// System API/DSM/API/bds_dsm_getErrors_DTC
///This function is used to get all DTCs with the specified status.
///
///=======
/// Remarks:
///=======
///    + The |GVL_dsm| is given for usage of defines.
///	
///----------
/// FFI:
///----------
///This API can be used in trusted partitions only. See Freedom from Interference (FFI) concept for more details.
///
///==================================================================		  			===================================================================================================
///Return value    								  									Description
///==================================================================		  			===================================================================================================
///16#0000: BDS_DSM_NO_ERROR_DU16														Got all DTC with specified status.
///16#0004: BDS_DSM_INVALID_PTR_DU16													Invalid Pointer.
///16#0005: BDS_DSM_MASK_ERROR_DU16													Invalid Mask.
///16#0007: BDS_DSM_INVALID_MAX_ERROR_DU16 											Invalid Max number of errors.
///16#0008:BDS_DSM_OVERFLOW_ERROR_DU16													Number of error are more than Max Error. 
///
///==================================================================		   			===================================================================================================
///
///
///=======
///Code Example:
///=======
///============================================================================
///
///PROGRAM DSM
///
///VAR
///
///	mask_s : UINT := BDS_DSM_SET_ACTIVE_ERROR_MASK_DU16;
///
///	startFromBegin_l: BOOL := TRUE;
///
///	maxNum_u16:UINT := 32;
///
///	error_count_u16: UINT;
///
///	dtc_u16: ARRAY [1..32] OF UINT;
///
///	status_u16: UINT;
///
///END_VAR
///
///
///(*Get errors*)
///
///status_u16 := bds_dsm_getErrors(mask_s,startFromBegin_l,maxNum_u16,ADR(error_count_u16),ADR(dtc_u16)); 
///
///IF status_u16 = BDS_DSM_NO_ERROR_DU16 THEN
///
///	(*Number of Errors has been read successfully*)
///
///END_IF
///
///============================================================================
///
{attribute 'external_name' := 'cmp_rts_bds_dsm_getErrors_DTC'}
FUNCTION bds_dsm_getErrors_DTC : UINT
VAR_INPUT
	///The kind of error status can be specified in detail by means of this mask.
	///
	///Possible values:
	///    + BDS_DSM_SET_ACTIVE_ERROR_MASK_DU16 ( 16#18 ) - Fault is active.
	///    + BDS_DSM_SET_TESTED_ONCE_MASK_DU16 ( 16#08 ) - DFC was tested at least once since start or reset.
	///    + BDS_DSM_SET_TESTED_OK_MASK_DU16 ( 16#20 ) - DFC was at least once ok tested since start or reset.  
	///    + BDS_DSM_SET_FAILED_SINCE_CLEAR_MASK_DU16 ( 16#80 ) - Fault occured at least once since error was deleted from memory.
	mask_s: UINT;
	///
	///    + TRUE: Query is started from the beginning of DFES.
	///    + FALSE: Query is continued with the next index where the last query was finished.
	startFromBegin_l: BOOL;
	///Maximal number of errors/DTCs which can be returned.
	maxNum_u16: UINT;
	///Pointer to a variable where the number of errors/DTCs is returned.
	num_pu16: POINTER TO UINT;
	///Pointer to a variable used to store DTC value.
	dtc_pu16: POINTER TO UINT;
END_VAR

END_FUNCTION

// System API/DSM/API/bds_dsm_getFIdPermission
///This function is used to get the permission of error reaction.
///
///=======
/// Remarks:
///=======
///    + The |GVL_dsm| is given for usage of defines.
///	
///----------
/// FFI:
///----------
///This API can be used in trusted partitions only. See Freedom from Interference (FFI) concept for more details.
///
///==================================================================		  			===================================================================================================
///Return value    								  									Description
///==================================================================		  			===================================================================================================
///TRUE																				Function has running permission.
///FALSE																				Function is blocked.
///
///==================================================================		   			===================================================================================================
///
///
///=======
///Code Example:
///=======
///============================================================================
///
///PROGRAM DSM
///
///VAR
///
///	fid_test:bds_dsm_fid_ts; 
///
///	result:bool;
///
///END_VAR
///
///
///fid_test.id := 001;
///
///(*Get the permission for FId*)
///
///result := bds_dsm_getFIdPermission(fid_test);
///
///============================================================================
///
{attribute 'external_name' := 'cmp_rts_bds_dsm_getFIdPermission'}
FUNCTION bds_dsm_getFIdPermission : BOOL
VAR_INPUT
	///Function Identifier (function or part of a function which is to be enabled or inhibited) : It is configured using easyConfig tool.
	fid_s: bds_dsm_fid_ts;
END_VAR

END_FUNCTION

// System API/DSM/API/Macro Functions/bds_dsm_DFC_fl
///It returns the fault level bit fields from DFC status word
{attribute 'external_name' := 'cmp_rts_bds_dsm_DFC_fl'}
FUNCTION bds_dsm_DFC_fl : USINT
VAR_INPUT
	dfc_u16: UINT;
END_VAR

END_FUNCTION

// System API/DSM/API/bds_dsm_getNumErrors
///This function returns the number of errors and the type of the errors is specified by a mask.
///
///=======
/// Remarks:
///=======
///    + The |GVL_dsm| is given for usage of defines.
///
///----------
/// FFI:
///----------
///This API can be used in trusted partitions . For untrusted partitions use |bds_dsm_getNumErrors_ffi|. See Freedom from Interference (FFI) concept for more details.
///	
///==================================================================		  			===================================================================================================
///Return value    								  									Description
///==================================================================		  			===================================================================================================
///16#0000: BDS_DSM_NO_ERROR_DU16														Update Number of Error is Successful.
///16#0004: BDS_DSM_INVALID_PTR_DU16													Invalid Pointer.
///16#0005: BDS_DSM_MASK_ERROR_DU16													Invalid Mask.
///16#000C: BDS_DSM_FFI_ACCESS_ERROR_DU16												Invalid Access to FFI variant API call.
///
///==================================================================		   			===================================================================================================
///
///
///=======
///Code Example:
///=======
///============================================================================
///
///PROGRAM DSM
///
///VAR
///
///	status_u16: UINT;
///
///	num_error_u16: UINT;
///
///END_VAR
///
///(*Get number of errors*)
///
///status_u16 := bds_dsm_getNumErrors(BDS_DSM_SET_ACTIVE_ERROR_MASK_DU16,ADR(num_error_u16));
///
///IF status_u16 = BDS_DSM_NO_ERROR_DU16 THEN
///
///	(*Number of Errors has been read successfully*)
///
///END_IF
///
///============================================================================
///
{attribute 'external_name' := 'cmp_rts_bds_dsm_getNumErrors'}
FUNCTION bds_dsm_getNumErrors : UINT
VAR_INPUT
	///The kind of error status can be specified in detail by means of this mask.
	///
	///Possible values:
	///    + BDS_DSM_SET_ACTIVE_ERROR_MASK_DU16 ( 16#18 ) - Fault is active.
	///    + BDS_DSM_SET_TESTED_ONCE_MASK_DU16 ( 16#08 ) - DFC was tested at least once since start or reset.
	///    + BDS_DSM_SET_TESTED_OK_MASK_DU16 ( 16#20 ) - DFC was at least once ok tested since start or reset.  
	///    + BDS_DSM_SET_FAILED_SINCE_CLEAR_MASK_DU16 ( 16#80 ) - Fault occured at least once since error was deleted from memory.
	mask_s: UINT;
	///Pointer to a variable where the number of errors/DFCs are returned.
	number_pu16: POINTER TO UINT;
END_VAR

END_FUNCTION

// System API/DSM/FFI_API/bds_dsm_getNumErrors_ffi
{attribute 'external_name' := 'cmp_rts_bds_dsm_getNumErrors_ffi'}
FUNCTION bds_dsm_getNumErrors_ffi : UINT
VAR_INPUT
	///The kind of error status can be specified in detail by means of this mask.
	///
	///Possible values:
	///    + BDS_DSM_SET_ACTIVE_ERROR_MASK_DU16 ( 16#18 ) - Fault is active.
	///    + BDS_DSM_SET_TESTED_ONCE_MASK_DU16 ( 16#08 ) - DFC was tested at least once since start or reset.
	///    + BDS_DSM_SET_TESTED_OK_MASK_DU16 ( 16#20 ) - DFC was at least once ok tested since start or reset.  
	///    + BDS_DSM_SET_FAILED_SINCE_CLEAR_MASK_DU16 ( 16#80 ) - Fault occured at least once since error was deleted from memory.
	mask_s: UINT;
	///Pointer to a variable where the number of errors/DFCs are returned.
	number_pu16: POINTER TO UINT;
END_VAR

END_FUNCTION

// System API/DSM/API/bds_dsm_getNumErrorsJ1939
///This functions returns the number of errors and the type of the errors is specified by a state and which were configured for J1939 only.
///
///=======
/// Remarks:
///=======
///    + The |GVL_dsm| is given for usage of defines.
///	+ Suspect Parameter Number (SPN), Failure Mode Identifier (FMI) and Lamp States can be configured in easyConfig.
///
///----------
/// FFI:
///----------
///This API can be used in trusted partitions only. See Freedom from Interference (FFI) concept for more details.
///
///-----
/// NOTICE:
///-----
///	+ SPN or FMI should be non zero to be visible in J1939.
///	
///==================================================================		  			===================================================================================================
///Return value    								  									Description
///==================================================================		  			===================================================================================================
///16#0000: BDS_DSM_NO_ERROR_DU16														Update Number of Error is Successful .
///16#0004: BDS_DSM_INVALID_PTR_DU16													Invalid Pointer.
///16#0005: BDS_DSM_STATE_ERROR_DU16													Invalid State.
///16#000A: BDS_DSM_WRONG_BUFFERSIZE_DU16												Buffersize is invalid.
///16#000B:BDS_DSM_NO_DTC_AVAILABLE_DU16												No more DTC is available.
///
///==================================================================		   			===================================================================================================
///
///
///=======
///Code Example:
///=======
///============================================================================
///
///PROGRAM DSM
///
///VAR
///
///	status_u16: UINT;
///
///	num_error_u16: UINT;
///
///END_VAR
///
///(*Get number of errors*)
///
///status_u16 := bds_dsm_getNumErrorsJ1939(ACTIVE_ERRORS,ADR(num_error_u16));
///
///IF status_u16 = BDS_DSM_NO_ERROR_DU16 THEN
///
///	(*Number of Errors has been read successfully*)
///
///END_IF
///
///============================================================================
///
{attribute 'external_name' := 'cmp_rts_bds_dsm_getNumErrorsJ1939'}
FUNCTION bds_dsm_getNumErrorsJ1939 : UINT
VAR_INPUT
	///The kind of error status can be specified in detail by means of this mask.
	///	+ ACTIVE_ERRORS(0)                      - Fault is Active.
	///	+ PREVIOUSLY_ACTIVE_ERRORS(1) - Fault was Previously Active.
	state_e: bds_dsm_state_te;
	///Pointer to a variable where the number of errors/DFCs are returned.
	number_pu8: POINTER TO USINT;
END_VAR

END_FUNCTION

// System API/DSM/API/Macro Functions/bds_dsm_DFC_fsc
///It returns the fault since clear bit fields from DFC status word
{attribute 'external_name' := 'cmp_rts_bds_dsm_DFC_fsc'}
FUNCTION bds_dsm_DFC_fsc : USINT
VAR_INPUT
	dfc_u16: UINT;
END_VAR

END_FUNCTION

// System API/DSM/API/bds_dsm_testError
///This function is used to check the status of a DFC.
///
///=======
/// Remarks:
///=======
///    + The |GVL_dsm| is given for usage of defines.
///
///----------
/// FFI:
///----------
///This API can be used in trusted partitions only. See Freedom from Interference (FFI) concept for more details.
///
///-----
/// NOTICE:
///-----
///	+ SPN or FMI should be non zero to be visible in J1939.
///	
///==================================================================		  			===================================================================================================
///Return value    								  									Description
///==================================================================		  			===================================================================================================
///16#0000: BDS_DSM_NO_ERROR_DU16														Update of Error status is successful.
///16#0001: BDS_DSM_DFC_ERROR_DU16														Invalid DFC.
///16#0004: BDS_DSM_INVALID_PTR_DU16													Invalid pointer.
///
///==================================================================		   			===================================================================================================
///
///
///=======
///Code Example:
///=======
///============================================================================
///
///PROGRAM DSM
///
///VAR
///
///	dfc_s: bds_dsm_dfc_ts;	
///
///	dfc_ts : DFC_bds_NoDebFault1;
///
///	status_dfc_u16:UINT;
///
///	result_u16: POINTER TO UINT;
///
///	status_u16: UINT;
///
///END_VAR
///
///(*To get the status of DFC*)
///
///dfc_s.id := dfc_ts.DFCid;
///
///status_u16 := bds_dsm_testError(dfc_s, ADR(status_dfc_u16)); 
///
///IF status_u16 = BDS_DSM_NO_ERROR_DU16 THEN
///
///	(*Status have been updated successfully*)
///
///END_IF
///
///============================================================================
///
{attribute 'external_name' := 'cmp_rts_bds_dsm_testError'}
FUNCTION bds_dsm_testError : UINT
VAR_INPUT
	///DFC name (identifier) : It is configured using easyConfig tool.
	dfc_s: bds_dsm_dfc_ts;
	///Pointer to a variable where the test result is returned. result is bit-coded.
	///
	///	+ 00:  ACTIVE_DFC_STATUS_DU8 (16#18) - Fault is active.
	///	+ 01:  TESTED_ONCE_STATUS_DU8 (16#08) - DFC was tested at least once since start or reset. 
	///	+ 10:  TESTED_OK_SINCE_CLEAR_DU8 (16#20) - DFC was at least once ok tested since start or reset.
	///	+ 11:   FAULT_SINCE_CLEAR_DU8 (16#80) - Fault occured at least once since error memory was deleted.
	result_u16: POINTER TO UINT;
END_VAR

END_FUNCTION

// System API/DSM/API/bds_dsm_test_ErrorDFC
///This function is used to check whether given DFC is Active , previously Active or Deactive .
///
///=======
/// Remarks:
///=======
///    + The |GVL_dsm| is given for usage of defines.
///	+ Status of the DFC is bit coded and the definition of each bit is given below.
///
///	
///----------
/// FFI:
///----------
///This API can be used in trusted partitions only. See Freedom from Interference (FFI) concept for more details.
///
///==================================================================		  			===================================================================================================
///Return value    								  									Description
///==================================================================		  			===================================================================================================
///16#0000: BDS_DSM_NO_ERROR_DU16														Update of Error is Successful .
///16#0001: BDS_DSM_DFC_ERROR_DU16														Invalid DFC.
///16#0004: BDS_DSM_INVALID_PTR_DU16													Invalid Pointer.
///
///==================================================================		   			===================================================================================================
///
///
///=======
///Code Example:
///=======
///============================================================================
///
///PROGRAM DSM
///
///VAR
///
///	dfc_s: bds_dsm_dfc_ts;	
///
///	dfc_ts : DFC_bds_NoDebFault1;
///
///	status_u8:USINT;
///
///	error_u16: UINT;
///
///END_VAR
///
///(*To get the status of DFC*)
///
///dfc_s.id := dfc_ts.DFCid;
///
///error_u16 := bds_dsm_test_ErrorDFC(dfc_s,ADR(status_u8));
///
///IF error_u16 = BDS_DSM_NO_ERROR_DU16 THEN
///
///	(*Error Status has been reported succesfully*)
///
///END_IF
///
///============================================================================
///
{attribute 'external_name' := 'cmp_rts_bds_dsm_test_ErrorDFC'}
FUNCTION bds_dsm_test_ErrorDFC : UINT
VAR_INPUT
	///DFC name (identifier) : It is configured using easyConfig tool.
	dfc_s: bds_dsm_dfc_ts;
	///Pointer to a variable where the test result is returned. result is bit-coded.
	///	+ BDS_DSM_STATUS_ACTIVE_MASK_DU8(16#01)             : 0th bit is set when error is active.
	///	+ BDS_DSM_STATUS_PREVIOUSLY_ACTIVE_MASK_DU8(16#02)  : 1st bit is set when error is previously active.
	///	+ BDS_DSM_STATUS_DEACTIVE_MASK_DU8(16#04)           : 2nd bit is set when error is deactivated.
	///	+ BDS_DSM_STATUS_TESTED_SINCE_CLEAR_MASK_DU8(16#08) : 3rd bit is set when error is tested since clear.
	///	+ BDS_DSM_STATUS_FAULT_SINCE_CLEAR_MASK_DU8(16#10)  : 4th bit is set when error is fault since clear.
	result_u8: POINTER TO USINT;
END_VAR

END_FUNCTION

// System API/DSM/API/bds_dsm_test_ErrorDTC
///This function is used to check whether given DTC is Active, Previously Active or Deactive .
///
///=======
/// Remarks:
///=======
///    + The |GVL_dsm| is given for usage of defines.
///
///	
///----------
/// FFI:
///----------
///This API can be used in trusted partitions only. See Freedom from Interference (FFI) concept for more details.
///
///==================================================================		  			===================================================================================================
///Return value    								  									Description
///==================================================================		  			===================================================================================================
///16#0000: BDS_DSM_NO_ERROR_DU16														Update of status is successful .
///16#0004: BDS_DSM_INVALID_PTR_DU16													Invalid Pointer.
///16#000B: BDS_DSM_NO_DTC_AVAILABLE_DU16 												Invalid DTC input.
///
///==================================================================		   			===================================================================================================
///
///
///=======
///Code Example:
///=======
///============================================================================
///
///PROGRAM DSM
///
///VAR
///
///	dfc_s: bds_dsm_dfc_ts;	
///
///	dfc_ts : DFC_bds_NoDebFault1;
///
///	status_u8:USINT;
///
///	error_u16: UINT;
///
///END_VAR
///
///(*To get the status of DTC*)
///
///dfc_s.id := dfc_ts.DFCid;
///
///error_u16 := bds_dsm_test_ErrorDTC(dfc_ts.DTC,ADR(status_u8));
///
///IF error_u16 = BDS_DSM_NO_ERROR_DU16 THEN
///
///	(*Error Status has been reported succesfully*)
///
///END_IF
///
///============================================================================
///
{attribute 'external_name' := 'cmp_rts_bds_dsm_test_ErrorDTC'}
FUNCTION bds_dsm_test_ErrorDTC : UINT
VAR_INPUT
	///DTC Value : It is configured using easyConfig tool.
	dtc_u16: UINT;
	///Pointer to a variable where the test result is returned. result is bit-coded.
	///	+ BDS_DSM_STATUS_ACTIVE_MASK_DU8(16#01)             : 0th bit is set when error is active.
	///	+ BDS_DSM_STATUS_PREVIOUSLY_ACTIVE_MASK_DU8(16#02)  : 1st bit is set when error is previously active.
	///	+ BDS_DSM_STATUS_DEACTIVE_MASK_DU8(16#04)           : 2nd bit is set when error is deactivated.
	///	+ BDS_DSM_STATUS_TESTED_SINCE_CLEAR_MASK_DU8(16#08) : 3rd bit is set when error is tested since clear.
	///	+ BDS_DSM_STATUS_FAULT_SINCE_CLEAR_MASK_DU8(16#10)  : 4th bit is set when error is fault since clear.
	result_u8: POINTER TO USINT;
END_VAR

END_FUNCTION

// System API/DSM/API/bds_dsm_updateDebError
///This function is used to update the DFCs configured with debouncing.
///
///=======
/// Remarks:
///=======
///    + The |GVL_dsm| is given for usage of defines.
///
///	
///----------
/// FFI:
///----------
///This API can be used in trusted partitions only. See Freedom from Interference (FFI) concept for more details.
///
///==================================================================		  			===================================================================================================
///Return value    								  									Description
///==================================================================		  			===================================================================================================
///16#0000: BDS_DSM_NO_ERROR_DU16														Update of Error is Successful.
///16#0001: BDS_DSM_DFC_ERROR_DU16														Invalid DFC.
///16#0002: BDS_DSM_DEBOUNCE_ERROR_DU16												Invalid Debounce method.
///16#0003: BDS_DSM_FAULT_PERCENT_ERROR_DU16											Invalid Error Percentage.
///
///==================================================================		   			===================================================================================================
///
///
///=======
///Code Example:
///=======
///============================================================================
///
///PROGRAM DSM
///
///VAR
///
///	dfc_s: bds_dsm_dfc_ts;	
///
///	dfc_ts : DFC_bds_NoDebFault1;
///
///	result_u16:UINT;
///
///	status_u16: UINT;
///	
///	tDiff_u32: UDINT;
///
///END_VAR
///
///(*Reporting the Error(debounce) with 100 percent fault percentage*)
///
///dfc_s.id := dfc_ts.DFCid;
///
///status_u16:=bds_dsm_updateDebError(dfc_s,result_u16,tDiff_u32);
///
///IF status_u16 = BDS_DSM_NO_ERROR_DU16 THEN
///
///	(*Error has been reported succesfully*)
///
///END_IF
///
///============================================================================
///
{attribute 'external_name' := 'cmp_rts_bds_dsm_updateDebError'}
FUNCTION bds_dsm_updateDebError : UINT
VAR_INPUT
	///DFC name (identifier) : It is configured using easyConfig tool.
	dfc_s: bds_dsm_dfc_ts;
	///Result of the check.
	///    + BDS_DSM_FAULT_PERCENT_00_DU8    : ok
	///    + BDS_DSM_FAULT_PERCENT_100_DU8  : not ok
	result_u16: UINT;
	///Time difference since last call in µs.
	///It is needed for time debounce types only. Please use 0 for other debounce types (e.g. event debounce types).    
	tDiff_u32: UDINT;
END_VAR

END_FUNCTION

// System API/DSM/API/bds_dsm_updateError
///This function is used to update DFCs configured with no debouncing. 
///
///=======
/// Remarks:
///=======
///    + The |GVL_dsm| is given for usage of defines.
///
///	
///----------
/// FFI:
///----------
///This API can be used in trusted partitions . For untrusted partitions use |bds_dsm_updateError_ffi|. See Freedom from Interference (FFI) concept for more details.
///
///==================================================================		  			===================================================================================================
///Return value    								  									Description
///==================================================================		  			===================================================================================================
///16#0000: BDS_DSM_NO_ERROR_DU16														Error is updated successfully.
///16#0001: BDS_DSM_DFC_ERROR_DU16														Invalid DFC.
///16#0002: BDS_DSM_DEBOUNCE_ERROR_DU16												Invalid Debounce method.
///16#0003: BDS_DSM_FAULT_PERCENT_ERROR_DU16											Invalid Error Percentage.
///16#000C: BDS_DSM_FFI_ACCESS_ERROR_DU16												Invalid Access to FFI variant API call.
///
///==================================================================		   			===================================================================================================
///=======
///Code Example:
///=======
///============================================================================
///
///PROGRAM DSM
///
///VAR
///
///	dfc_s: bds_dsm_dfc_ts;	
///
///	dfc_ts : DFC_bds_NoDebFault1;
///
///	result_u16:UINT;
///
///	status_u16: UINT;
///	
///	tDiff_u32: UDINT;
///
///END_VAR
///
///(*Reporting the Error(debounce) with 100 percent fault percentage*)
///
///dfc_s.id := dfc_ts.DFCid;
///
///status_u16 := bds_dsm_updateError(dfc_s,BDS_DSM_FAULT_PERCENT_100_DU8); 
///
///IF status_u16 = BDS_DSM_NO_ERROR_DU16 THEN
///
///	(*Error has been reported succesfully*)
///
///END_IF
///
///============================================================================
///
{attribute 'external_name' := 'cmp_rts_bds_dsm_updateError'}
FUNCTION bds_dsm_updateError : UINT
VAR_INPUT
	///DFC name (identifier) : It is configured using easyConfig tool.
	dfc_s: bds_dsm_dfc_ts;
	///Result of the check.
	///    + BDS_DSM_FAULT_PERCENT_00_DU8   : ok
	///    + BDS_DSM_FAULT_PERCENT_100_DU8 : not ok
	result_u16: UINT;
END_VAR

END_FUNCTION

// System API/DSM/FFI_API/bds_dsm_updateError_ffi
{attribute 'external_name' := 'cmp_rts_bds_dsm_updateError_ffi'}
FUNCTION bds_dsm_updateError_ffi : UINT
VAR_INPUT
	///DFC name (identifier) : It is configured using easyConfig tool.
	dfc_s: bds_dsm_dfc_ts;
	///Result of the check.
	///    + BDS_DSM_FAULT_PERCENT_00_DU8   : ok
	///    + BDS_DSM_FAULT_PERCENT_100_DU8 : not ok
	result_u16: UINT;
END_VAR

END_FUNCTION

// System API/DSM/API/Macro Functions/bds_dsm_DFC_ms
///It returns the memory status bit fields from DFC status word
{attribute 'external_name' := 'cmp_rts_bds_dsm_DFC_ms'}
FUNCTION bds_dsm_DFC_ms : USINT
VAR_INPUT
	dfc_u16: UINT;
END_VAR

END_FUNCTION

// System API/DSM/API/bds_dsm_updateError_DTC
///This function is used to update DFES entry, with the help of DTC.
///
///=======
/// Remarks:
///=======
///    + The |GVL_dsm| is given for usage of defines.
///
///	
///----------
/// FFI:
///----------
///This API can be used in trusted partitions only. See Freedom from Interference (FFI) concept for more details.
///
///==================================================================		  			===================================================================================================
///Return value    								  									Description
///==================================================================		  			===================================================================================================
///16#0000: BDS_DSM_NO_ERROR_DU16														Error is updated successfully.
///16#0002: BDS_DSM_DEBOUNCE_ERROR_DU16												Invalid Debounce method.
///16#0003: BDS_DSM_FAULT_PERCENT_ERROR_DU16											Invalid Error Percentage.
///16#000B: BDS_DSM_NO_DTC_AVAILABLE_DU16												Invalid DTC.
///
///==================================================================		   			===================================================================================================
///
///
///=======
///Code Example:
///=======
///============================================================================
///
///PROGRAM DSM
///
///VAR
///
///	dfc_s: bds_dsm_dfc_ts;	
///
///	dfc_ts : DFC_bds_NoDebFault1;
///
///	result_u16:UINT;
///
///	status_u16: UINT;
///	
///	tDiff_u32: UDINT;
///
///END_VAR
///
///(*Reporting the Error(debounce) with 100 percent fault percentage*)
///
///dfc_s.id := dfc_ts.DFCid;
///
///status_u16 :=bds_dsm_updateError_DTC(dfc_ts.DTC, result_u16, tDiff_u32); 
///
///IF status_u16 = BDS_DSM_NO_ERROR_DU16 THEN
///
///	(*Error has been reported succesfully*)
///
///END_IF
///
///============================================================================
{attribute 'external_name' := 'cmp_rts_bds_dsm_updateError_DTC'}
FUNCTION bds_dsm_updateError_DTC : UINT
VAR_INPUT
	///DTC value : It is configured using easyConfig tool.
	dtc_u16: UINT;
	///Result of the check,
	///    + BDS_DSM_FAULT_PERCENT_00_DU8     : ok,
	///    + BDS_DSM_FAULT_PERCENT_100_DU8   : not ok.
	result_u16: UINT;
	///Time difference since last call in µsec.
	tdiff_u32: UDINT;
END_VAR

END_FUNCTION

// System API/DSM/API/Macro Functions/bds_dsm_DFC_t
///It returns the test status bit fields from DFC status word
{attribute 'external_name' := 'cmp_rts_bds_dsm_DFC_t'}
FUNCTION bds_dsm_DFC_t : USINT
VAR_INPUT
	dfc_u16: UINT;
END_VAR

END_FUNCTION

// System API/DSM/API/Macro Functions/bds_dsm_DFC_tf
///It returns the test finalized bit fields from DFC status word
{attribute 'external_name' := 'cmp_rts_bds_dsm_DFC_tf'}
FUNCTION bds_dsm_DFC_tf : USINT
VAR_INPUT
	dfc_u16: UINT;
END_VAR

END_FUNCTION

// System API/DSM/API/Macro Functions/bds_dsm_DFC_tsc
///It returns the test since clear bit fields from DFC status word
{attribute 'external_name' := 'cmp_rts_bds_dsm_DFC_tsc'}
FUNCTION bds_dsm_DFC_tsc : USINT
VAR_INPUT
	dfc_u16: UINT;
END_VAR

END_FUNCTION

// I/O API/IN legacy/API/bds_in_ai
///Provides the ADC (analog to digital converter) voltage of the input in digits.
///
///=======
/// Remarks:
///=======
///    + The raw value  in digits ranges from  0 to 25000 with the resolution of 200µV per digit for 0 to 5V inputs. For other ranges the resolution will vary accordingly as shown below.
///
///----------
/// FFI:
///----------
///This API can be used in trusted partitions only. See Freedom from Interference (FFI) concept for more details.
///
///==================================================================		  			===================================================================================================
///Voltage range    								  									Per digit resolution
///==================================================================		  			===================================================================================================
///0 - 5V																				200
///0- 20V																				800
///0-32V																				1600
///0-40V																				1240
///
///==================================================================		   			===================================================================================================
///
///
///==================================================================		  			===================================================================================================
///Return value    								  									Description
///==================================================================		  			===================================================================================================
///0																					No error
///1																					Invalid parameter
///2																					Function call was erroneous
///
///==================================================================		   			===================================================================================================
///
///=======
///Code Example:
///=======
///============================================================================
///
///PROGRAM appl_10ms_task
///  VAR
///  
///    digitsK59_u16: UINT := 16#00;
///  END_VAR
///
///  (* get the ADC value of input K59 *)
///
///  bds_in_ai(bds_in_aiv_signal_te.K59, ADR(digitsK59_u16))
///
///END
///
///============================================================================
{attribute 'external_name' := 'cmp_rts_bds_in_ai'}
FUNCTION bds_in_ai : USINT
VAR_INPUT
	///The signal name that is assigned to the respective pin configured as voltage input
	signal_e: UINT;
	///Storage address of the value.
	///
	///Range:
	///0 to 25000  [200µV] per digit
	value_pu16: POINTER TO UINT;
END_VAR

END_FUNCTION

// I/O API/IN legacy/API/bds_in_aic
///Provides the analog current of the input.
///
///=======
/// Remarks:
///=======
///    + The inputs support the reading of analog current if the shunt is activated using easyConfig (eC).
///    + The voltage drop across the shunt is measured with the parallel running analog voltage input. (see the INFO).
///    + The measurement range is 0 to 24000µA. 
///    + The shunt must be protected if the current exceeds 23500µA. After the deactivation of the shunt, recovery time of 2s is required. 
///    + After the recovery time elapses, the shunt can be activated again with |bds_sys_do|.
///    + For more info about the shunt protection see  |bds_in_aic_getStatus|.
///
///----------
/// FFI:
///----------
///This API can be used in trusted partitions only. See Freedom from Interference (FFI) concept for more details.
///
///------
///INFO:
///------
///    + When DSM/AIC is selected in eC then it is not possible to select the voltage range and PullUp and  PullDown. These fields are greyed out.
///    + The PullUp and PullDown configuration is set to external (this corresponds to float) because to avoid the offset current provided by the PullUp or PullDown current strength.
///
///	
///==================================================================		  			===================================================================================================
///Return value    								  									Description
///==================================================================		  			===================================================================================================
///0																					No error
///1																					Invalid parameter
///2																					Function call was erroneous
///3																					Shunt not activated
///
///==================================================================		   			===================================================================================================
///
///=======
///Code Example:
///=======
///============================================================================
///
///PROGRAM appl_10ms_task
///  VAR
///  
///    uA_K54_u16: UINT := 16#00;
///  END_VAR
///
/// (* As a precondition K54_VI must be enabled for the current measurement,
///   means that the shunt at the input shall be activated (configured with eC) *)
///
/// (* get current value *)
///
///  bds_in_aic(bds_in_fi_signal_te.K54_VI, ADR(uA_K54_u16));
///END
///
///============================================================================
{attribute 'external_name' := 'cmp_rts_bds_in_aic'}
FUNCTION bds_in_aic : USINT
VAR_INPUT
	///The signal name that is assigned to the respective pin configured as current input
	signal_e: UINT;
	///Storage address of the value.
	///
	///Range:
	///0 to 24000 [µA]
	value_pu16: POINTER TO UINT;
END_VAR

END_FUNCTION

// System API/DSM/API/bds_dsm_getDFC_Status
///This function is used to get the 16 bit DFC status word of specified DFC.
///
///=======
/// Remarks:
///=======
///    + The |GVL_dsm| is given for usage of defines.
///	   + For information on 16 bit DFC status word refer Diagnostic Fault Check. 
///
///----------
/// FFI:
///----------
///This API can be used in trusted partitions . For untrusted partitions use |bds_dsm_getDFC_Status_ffi|. See Freedom from Interference (FFI) concept for more details.
///
///==================================================================		  			===================================================================================================
///Return value    								  									Description
///==================================================================		  			===================================================================================================
///16#0000: BDS_DSM_NO_ERROR_DU16														Update of Error is Successful .
///16#0001: BDS_DSM_DFC_ERROR_DU16														Invalid DFC.
///16#0004: BDS_DSM_INVALID_PTR_DU16													Invalid Pointer.
///16#000C: BDS_DSM_FFI_ACCESS_ERROR_DU16												Invalid Access to FFI variant API call.
///
///==================================================================		   			===================================================================================================
///
///
///=======
///Code Example:
///=======
///============================================================================
///
///PROGRAM BDS_DSM_getDFC_Status_TEST
///
///VAR
///
///	status_u16: UINT;
///
///	dfc_s: bds_dsm_dfc_ts;	
///
///	dfc_ts : DFC_bds_NoDebFault1;
///
///	error_u16:UINT;
///
///END_VAR
///
///dfc_s.id := dfc_ts.DFCid;
///
///(*Deletes the Error status from DFC and related DFES entry*)
///
///error_u16 := bds_dsm_getDFC_Status(dfc_s, ADR(status_u16));
///
///if error_u16 = BDS_DSM_NO_ERROR_DU16 THEN
///
///	(*Error Status has been reported succesfully*)
///
///END_IF
///
///============================================================================
///
{attribute 'external_name' := 'cmp_rts_bds_dsm_getDFC_Status'}
FUNCTION bds_dsm_getDFC_Status : UINT
VAR_INPUT
	///DFC name (identifier) : It is configured using easyConfig tool.
	dfc_s: bds_dsm_dfc_ts;
	///Pointer to variable where the 16 bit DFC status word is returned.
	dfc_status: POINTER TO UINT;
END_VAR

END_FUNCTION

// System API/DSM/FFI_API/bds_dsm_getDFC_Status_ffi
{attribute 'external_name' := 'cmp_rts_bds_dsm_getDFC_Status_ffi'}
FUNCTION bds_dsm_getDFC_Status_ffi : UINT
VAR_INPUT
	///DFC name (identifier) : It is configured using easyConfig tool.
	dfc_s: bds_dsm_dfc_ts;
	///Pointer to variable where the 16 bit DFC status word is returned.
	dfc_status: POINTER TO UINT;
END_VAR

END_FUNCTION

// System API/DSM/API/bds_dsm_getDFES
///This function is used to get the data of one or more DFES entries.
///
///=======
/// Remarks:
///=======
///    + The |GVL_dsm| is given for usage of defines.
///
///----------
/// FFI:
///----------
///This API can be used in trusted partitions only. See Freedom from Interference (FFI) concept for more details.
///
///-----
/// NOTICE:
///-----
///    + On a maximum, 32 different DFES entries are possible. 
///    + Status Mask will take time (max. 10ms) to update in global mask so return status has to be monitored.
///	
///==================================================================		  			===================================================================================================
///Return value    								  									Description
///==================================================================		  			===================================================================================================
///16#0000: BDS_DSM_NO_ERROR_DU16														Update Number of Error is successful .
///16#0004: BDS_DSM_INVALID_PTR_DU16													Invalid Pointer.
///16#0005: BDS_DSM_MASK_ERROR_DU16													Invalid Mask.
///16#0007: BDS_DSM_INVALID_MAX_ERROR_DU16 											Invalid Max Error.
///
///==================================================================		   			===================================================================================================
///
///
///=======
///Code Example:
///=======
///============================================================================
///
///PROGRAM BDS_DSM_getDFES_TEST
///
///VAR
///
///	mask_s : UINT := BDS_DSM_SET_ACTIVE_ERROR_MASK_DU16;
///
///	startFromBegin_l: BOOL := TRUE;
///
///	maxNum_u16:UINT := 32;
///
///	error_count_u16: UINT;
///
///	dfc_active_as: ARRAY [1..32] OF bds_dsm_dfc_ts;
///
///	status_u16: UINT;
///
///END_VAR
///
///dfc_s.id := dfc_ts.DFCid;
///
///(*Get DFES entries*)
///
///status_u16 := bds_dsm_getDFES(mask_s, TRUE, maxNum_u16, ADR(error_count_u16), ADR(dfc_active_as));
///
///if status_u16 = BDS_DSM_NO_ERROR_DU16 THEN
///
///	(*Numbers of Errors have been read successfully*)
///
///END_IF
///
///============================================================================
///
{attribute 'external_name' := 'cmp_rts_bds_dsm_getDFES'}
FUNCTION bds_dsm_getDFES : UINT
VAR_INPUT
	///The kind of error status can be specified in detail by means of this mask.
	///
	///Possible values:
	///    + BDS_DSM_SET_ACTIVE_ERROR_MASK_DU16 ( 16#18 ) - Fault is active.
	///    + BDS_DSM_SET_TESTED_ONCE_MASK_DU16 ( 16#08 ) - DFC was tested at least once since start or reset.
	///    + BDS_DSM_SET_TESTED_OK_MASK_DU16 ( 16#20 ) - DFC was at least once ok tested since start or reset.  
	///    + BDS_DSM_SET_FAILED_SINCE_CLEAR_MASK_DU16 ( 16#80 ) - Fault occured at least once since error was deleted from memory.
	mask_s: UINT;
	///TRUE: Query is started from the beginning of DFES.
	startFromBegin_l: BOOL;
	///Maximal number of errors/DFCs is returned. The BSW will return at max. 32 values (the max. size of DFES).
	maxNum_u16: UINT;
	///Pointer to a variable where the number of errors/DFC's is returned.
	num_pu16: POINTER TO UINT;
	///Pointer to all data of a DFES entry.
	data_pas: POINTER TO bds_dfes_ts;
END_VAR

END_FUNCTION

// I/O API/IN legacy/API/bds_in_ri_getTemp
///Provides the temperature value.
///
///=======
/// Remarks:
///=======
///   + The measurement range of the supported BSW sensors are from -50 to150°C with a resolution of 1°C, for more information see |bds_in_ri_cfgTemp|.
///   + If the resistance value is higher than 65535 ohm a value of 333°C is indicated as an invalid temperature.
///   
///
///----------
/// FFI:
///----------
///This API can be used in trusted partitions only. See Freedom from Interference (FFI) concept for more details.
///   
///==================================================================		  			===================================================================================================
///Return value    								  									Description
///==================================================================		  			===================================================================================================
///0																					No error
///1																					Invalid parameter
///2																					Resistance is out of range
///
///==================================================================		   			===================================================================================================
///
///=======
///Code Example:
///=======
///============================================================================
///
///PROGRAM PLC_PRG
///
///	VAR
///	
///		tempK60_s16: INT := 16#00;
///		
///		tempK58_s16: INT := 16#00;
///			
///		Init_flag_u8:USINT:=0;
///	
///	END_VAR
///  
///IF(Init_flag_u8=0) THEN (*To make api call once in application*)
///
///	(*get temperature of input K60 and K58*)
///	
///	bds_in_ri_getTemp(bds_in_ri_signal_te.K60, ADR(tempK60_s16));
///	
///	bds_in_ri_getTemp(bds_in_ri_signal_te.K58, ADR(tempK58_s16));
///	
///	Init_flag_u8:=1;
///  
///END_IF
///
///============================================================================
{attribute 'external_name' := 'cmp_rts_bds_in_ri_getTemp'}
FUNCTION bds_in_ri_getTemp : USINT
VAR_INPUT
	///The signal name that is assigned to the respective pin configured as resistance input
	signal_e: UINT;
	///Storage address OF the value.
	///
	///Range:
	///-50..150 [°C]
	value_s16: POINTER TO INT;
END_VAR

END_FUNCTION

// Communication API/ISOBUS/API/bds_isobus_cfgAddrClaimFormat
///This function configures the Address Claim Delay Format according to the J1939/ISOBUS standard.
///
///=======
/// Remarks:
///=======
///   + The use of this API is optional. By default the Address claim delay format is configured with ISOBUS standard.
///   + This function must be called once during the configuration of the ISOBUS communication stack before |bds_isobus_initComm| and |bds_isobus_setCaAddr|.
///   + According to the J1939-81 standard for the Source Address 0-127 and  248-253 ranges may omit the 250ms delay after the Address Claim Message is sent.
///   + According to the ISO 11783-5 standard for the complete Source Address range the 250ms delay to be used after the Address Claim Message is sent.
///   + The |GVL_isobus| is given for usage of defines.
///   + This function should be called only once in the application.
///
///----------
/// WARNING:
///----------
///
///This function should be called only once in the application.
///
///----------
/// FFI:
///----------
///This API can be used in trusted partitions only. See Freedom from Interference (FFI) concept for more details.
///
///==================================================================		  			===================================================================================================
///Return value    								  									Description
///==================================================================		  			===================================================================================================
///0: BDS_ISOBUS_RC_NO_ERRORS_DU16														Function was executed without errors.
///22: BDS_ISOBUS_RC_CFG_NOTALLOWED_DU16												Function must be called before |bds_isobus_initComm|, but it was called afterwards.
///
///==================================================================		   			===================================================================================================
///
///=======
///Code Example:
///=======
///============================================================================
///
///This Api should be called only once in application.
///
///
///PROGRAM Isobus_prg
///
///VAR
///
///    Flag_u8:USINT:=0;
///	
///    retval_u16: UINT;
///	
///END_VAR
///
///(*call the api once*)
///
///IF(Flag_u8=0)THEN
///    
///    (*configure the Address Claim Delay Format acc. to the ISOBUS standard*)
///	
///    retval_u16:=bds_isobus_cfgAddrClaimFormat(FALSE);
///        
///    (*define the controller application name, required for address claiming*)
///	
///    bds_isobus_setCaName(1,16#00,16#02,16#00,16#01,16#81,16#01,16#01,16#33,BDS_ISOBUS_OWN_SN_DU32);
///    
///    (*define the initial source address and the CAN channel for the CA instance 1*)
///	
///    bds_isobus_setCaAddr(1,BDS_CAN_3_D,16#10);
///    
///    (*initialize and start isobus communication for all instances on this CAN channel*)
///	
///    bds_isobus_initComm(bds_can_Chnl_te.BDS_CAN_3_D, 50);
///	
///    Flag_u8:=1;
///    
///END_IF
///
///============================================================================
{attribute 'external_name' := 'cmp_rts_bds_isobus_cfgAddrClaimFormat'}
FUNCTION bds_isobus_cfgAddrClaimFormat : UINT
VAR_INPUT
	///Format of the Address Claim Delay.
	///
	///Possible values:
	///   + TRUE = Address Claim Delay according to J1939.
	///   + FALSE = Address Claim Delay according to ISOBUS.
	j1939Format_l: BOOL;
END_VAR

END_FUNCTION

// Communication API/ISOBUS/API/bds_isobus_initComm
///This function configures and starts the ISOBUS communication stack for all instances on one CAN channel.
///
///=======
/// Remarks:
///=======
///   + This function must be called once per CAN channel for the start of all instances of the ISOBUS communication stack on this CAN channel.
///   + After the initialization an Address Claim procedure will be started. This means that all instances on the corresponding CAN channel will send an AddressClaim message.
///   + If the same CAN bus is also used for further communication, ensure that the CAN IDs are uniquely assigned.
///   + The parameter maxTime_u8 defines the maximum allowed run time of the ISOBUS task in %, related to the ISOBUS cycle time.
///   + The ISOBUS cycle time is 10ms.
///   + The ISOBUS cycle time can be changed to 1ms or 5ms from easyConfig.
///   + The |GVL_isobus| is given for usage of defines.
///   + This function should be called only once in the application.
///   
///----------
/// WARNING:
///----------
///
///This function should be called only once in the application.
///
///----------
/// FFI:
///----------
///This API can be used in trusted partitions only. See Freedom from Interference (FFI) concept for more details.
///
///==================================================================		  			===================================================================================================
///Return value    								  									Description
///==================================================================		  			===================================================================================================
///None.																				-
///
///==================================================================		   			===================================================================================================
///
///=======
///Code Example:
///=======
///============================================================================
///
///This Api should be called only once in application.
///
///PROGRAM Isobus_prg
///
///VAR
///
///    Flag_u8:USINT:=0;
///
///    EcuType_as8: ARRAY[1..200] OF STRING := ['Main ECU'];
///
///    EcuManu_as8: ARRAY[1..150] OF STRING := ['BOSCH REXROTH'];
///
///    ApplTask_as8: ARRAY[1..100] OF STRING := ['EHR'];    
///
///END_VAR
///
///(*call the api once*)
///
///IF(Flag_u8=0)THEN
///    
///    (* optionally define some ECU information of the controller application for the PGNs HW-ID and SW-ID: *)
///
///    bds_isobus_setCaInfo(2,16#0,ADR(EcuType_as8),ADR(EcuManu_as8),ADR(ApplTask_as8));
///        
///    (*define the controller application name, required for address claiming*)
///
///    bds_isobus_setCaName(1,16#00,16#02,16#00,16#01,16#81,16#01,16#01,16#33,BDS_ISOBUS_OWN_SN_DU32);
///    
///    (*define the initial source address and the CAN channel for the CA instance 1*)
///
///    bds_isobus_setCaAddr(1,BDS_CAN_3_D,16#10);
///    
///    (*initialize and start isobus communication for all instances on this CAN channel*)
///
///    bds_isobus_initComm(bds_can_Chnl_te.BDS_CAN_3_D, 50);
///    
///    Flag_u8:=1;
///    
///END_IF
///
///============================================================================
{attribute 'external_name' := 'cmp_rts_bds_isobus_initComm'}
FUNCTION bds_isobus_initComm : BOOL
VAR_INPUT
	///Indicates the CAN channel.
	///
	///Possible values for RC18-12/40, RC27-18/40:
	///   + BDS_CAN_1_D(0)
	///   + BDS_CAN_2_D(1)
	///   + BDS_CAN_3_D(2)
	///   + BDS_CAN_4_D(3)
	canChnl_e: bds_can_Chnl_te;
	///Maximum allowed run time of the isobus task, related to the ISOBUS cycle time:
	///
	///Value range: 1..99 %    (recommended: 20%).
	maxTime_u8: USINT;
END_VAR

END_FUNCTION

// Communication API/ISOBUS/API/bds_isobus_setCaInfo
///This function defines ECU information strings for the hardware and software identification of a controller application.
///
///=======
/// Remarks:
///=======
///   + This function can be called for each controller application with different string definitions.
///   + Each of the parameter strings may have a length of 200 characters but the total data length of the corresponding PGN will be truncated to 300 characters.
///   + The impact of this function on the contents of the PGN request answers of PGN 16#00FDC5 and 16#00FEDA is described here.
///   + The |GVL_isobus| is given for usage of defines.
///   + This function should be called only once in the application.
///
///----------
/// FFI:
///----------
///This API can be used in trusted partitions only. See Freedom from Interference (FFI) concept for more details.
///   
///==================================================================		  			===================================================================================================
///Return value    								  									Description
///==================================================================		  			===================================================================================================
///None.																				None.
///
///==================================================================		   			===================================================================================================
///
///=======
///Code Example:
///=======
///============================================================================
///
///This Api should be called only once in application.
///
///PROGRAM Isobus_prg
///
///VAR
///
///    Flag_u8:USINT:=0;
///	
///	(*Use the same Array size in the application*)
///	
///    EcuType_as8: ARRAY[1..20] OF STRING := ['Main ECU'];
///
///    EcuManu_as8: ARRAY[1..20] OF STRING := ['BOSCH REXROTH'];
///
///    ApplTask_as8: ARRAY[1..20] OF STRING := ['EHR'];    
///
///END_VAR
///
///(*call the api once*)
///
///IF(Flag_u8=0)THEN
///    
///    (* optionally define some ECU information of the controller application for the PGNs HW-ID and SW-ID: *)
///
///    bds_isobus_setCaInfo(2,16#0,ADR(EcuType_as8),ADR(EcuManu_as8),ADR(ApplTask_as8));
///        
///    (*define the controller application name, required for address claiming*)
///
///    bds_isobus_setCaName(1,16#00,16#02,16#00,16#01,16#81,16#01,16#01,16#33,BDS_ISOBUS_OWN_SN_DU32);
///    
///    (*define the initial source address and the CAN channel for the CA instance 1*)
///
///    bds_isobus_setCaAddr(1,BDS_CAN_3_D,16#10);
///    
///    (*initialize and start isobus communication for all instances on this CAN channel*)
///
///    bds_isobus_initComm(bds_can_Chnl_te.BDS_CAN_3_D, 50);
///    
///    Flag_u8:=1;
///    
///END_IF
///
///
///============================================================================
{attribute 'external_name' := 'cmp_rts_bds_isobus_setCaInfo'}
FUNCTION bds_isobus_setCaInfo : BOOL
VAR_INPUT
	///ISOBUS instance number. This number identifies one instance of the ISOBUS stack.
	///
	///Value range: 1..n
	///n is the number of ISOBUS instances configured by easyConfig. 
	instanceNum_u8: USINT;
	///Pointer to a character string with the ECU location or NULL pointer.
	///If a string was defined with this parameter then it will become a part of the response of the PGN request to PGN 16#00FDC5 (ECU identification information).
	///
	///The max. string length is 200 characters, but the total data length of the PGN 16#00FDC5 (ECU identification) is limited to 300 characters
	ecuLoc_pas8: POINTER TO ARRAY[1..200] OF STRING;
	///Pointer to a character string with the ECU type or NULL pointer.
	///If a string was defined with this parameter then it will become a part of the response of the PGN request to PGN 16#00FDC5 (ECU identification information).
	///
	///The max. string length is 200 characters, but the total data length of the PGN 16#00FDC5 (ECU identification) is limited to 300 characters.
	ecuType_pas8: POINTER TO ARRAY[1..200] OF STRING;
	///Pointer to a character string with the ECU manufacturer or NULL pointer.
	///If a string was defined with this parameter then it will become a part of the response of the PGN request to PGN 16#00FDC5 (ECU identification information).
	///
	///The max. string length is 200 characters, but the total data length of the PGN 16#00FDC5 (ECU identification) is limited to 300 characters.
	ecuMan_pas8: POINTER TO ARRAY[1..200] OF STRING;
	///Pointer to a character string with the application task name or NULL pointer.
	///If a string was defined with this parameter then it will become a part of the response of the PGN request to PGN 16#00FEDA (Software identification).
	///
	///The max. string length is 200 characters, but the total data length of the PGN 16#00FEDA (Software identification) is limited to 300 characters.
	applTask_pas8: POINTER TO ARRAY[1..200] OF STRING;
END_VAR

END_FUNCTION

// Communication API/ISOBUS/API/bds_isobus_setCaName
///This function defines the name of one controller application for the ISOBUS communication.
///
///=======
/// Remarks:
///=======
///   + The name is defined for one specific ISOBUS instance.
///   + The name may be changed later on with a further call of this function.
///   + The controller application (CA) name is mainly used for the Address Claim procedure during start up.
///   + Other controllers can ask for the CA name with a requestPGN for the PGN 16#EEFF (AddressClaimed).
///   + This function also defines the arbitrary address capability feature of the CA.
///   + The |GVL_isobus| is given for usage of defines.
///   + This function should be called only once in the application.
///
///----------
/// FFI:
///----------
///This API can be used in trusted partitions only. See Freedom from Interference (FFI) concept for more details.
///   
///==================================================================		  			===================================================================================================
///Return value    								  									Description
///==================================================================		  			===================================================================================================
///None.																				None.
///
///==================================================================		   			===================================================================================================
///
///=======
///Code Example:
///=======
///============================================================================
///
///This Api should be called only once in application.
///
///PROGRAM Isobus_prg
///
///VAR
///
///    Flag_u8:USINT:=0;
///
///    EcuType_as8: ARRAY[1..200] OF STRING := ['Main ECU'];
///
///    EcuManu_as8: ARRAY[1..150] OF STRING := ['BOSCH REXROTH'];
///
///    ApplTask_as8: ARRAY[1..100] OF STRING := ['EHR'];    
///
///END_VAR
///
///(*call the api once*)
///
///IF(Flag_u8=0)THEN
///    
///    (* optionally define some ECU information of the controller application for the PGNs HW-ID and SW-ID: *)
///
///    bds_isobus_setCaInfo(2,16#0,ADR(EcuType_as8),ADR(EcuManu_as8),ADR(ApplTask_as8));
///        
///    (*define the controller application name, required for address claiming*)
///
///    bds_isobus_setCaName(1,16#00,16#02,16#00,16#01,16#81,16#01,16#01,16#33,BDS_ISOBUS_OWN_SN_DU32);
///    
///    (*define the initial source address and the CAN channel for the CA instance 1*)
///
///    bds_isobus_setCaAddr(1,BDS_CAN_3_D,16#10);
///    
///    (*initialize and start isobus communication for all instances on this CAN channel*)
///
///    bds_isobus_initComm(bds_can_Chnl_te.BDS_CAN_3_D, 50);
///    
///    Flag_u8:=1;
///    
///END_IF
///
///
///============================================================================
{attribute 'external_name' := 'cmp_rts_bds_isobus_setCaName'}
FUNCTION bds_isobus_setCaName : BOOL
VAR_INPUT
	///ISOBUS instance number. This number identifies one instance of the ISOBUS stack.
	///
	///Value range: 1..n
	///n is the number of ISOBUS instances configured by easyConfig. 
	instanceNum_u8: USINT;
	///Arbitrary Address Capability (1 bit):
	///This bit defines whether the ISOBUS stack shall search for a new source address in case of an address conflict during the address claiming procedure.
	///
	///Value range: 0..1
	arbitAddrCapable_u8: USINT;
	///Industry group (3 bit):
	///
	///Value range: 0..7
	industryGroup_u8: USINT;
	///Device instance (4 bit):
	///
	///Value range: 0..15
	deviceInstance_u8: USINT;
	///Device class (7 bit):
	///
	///Value range: 0..127
	deviceClass_u8: USINT;
	///Function (8 bit):
	///
	///Value range: 0..255
	function_u8: USINT;
	///Function instance (5 bit):
	///
	///Value range: 0..32
	functionInstance_u8: USINT;
	///ECU instance (3 bit):
	///
	///Value range: 0..7
	ecuInstance_u8: USINT;
	///Manufacturer code (11 bit):
	///
	///Value range: 0..2047
	manufacturerCode_u16: UINT;
	///Serial number (21 bit):
	///
	///Value range: 0..16#1FFFFF  or  BDS_ISOBUS_OWN_SN_DU32 to use the lowest 21 bits of the ECU serial number
	serialNumber_u32: UDINT;
END_VAR

END_FUNCTION

// Communication API/ISOBUS/API/bds_isobus_setCaAddr
///This function defines the source address of one ISOBUS controller application and assignes it to a CAN channel.
///
///=======
/// Remarks:
///=======
///   + This function must be called for each new controller application before starting the communication on the corresponding CAN channel with the API function |bds_isobus_initComm|.
///   + The source address but not the CAN channel may be changed later on with a further call of this function.
///   + If the source will be changed with this function while the communication is already running then an address claim message will be sent with the new source address.
///   + The given source address is used within all transmitted messages, but this address may be changed within the Address Claim procedure.
///   + The currently active source address can be read with the API function |bds_isobus_getCaAddr|.
///   + The |GVL_isobus| is given for usage of defines.
///   + This function should be called only once in the application.
///
///----------
/// FFI:
///----------
///This API can be used in trusted partitions only. See Freedom from Interference (FFI) concept for more details.
///   
///==================================================================		  			===================================================================================================
///Return value    								  									Description
///==================================================================		  			===================================================================================================
///0: BDS_ISOBUS_RC_NO_ERRORS_DU16														Function was executed without errors.
///80: BDS_ISOBUS_RC_INV_INST_NUM_DU16													Invalid instance number.
///81: BDS_ISOBUS_RC_INV_CAN_CHNL_DU16													Invalid CAN channel.
///82: BDS_ISOBUS_RC_INV_CA_ADDR_DU16													Invalid own CA address (>253).
///83: BDS_ISOBUS_RC_CA_ADDR_IN_USE_DU16												The given own CA address is already in use by another CA on the same CAN channel. This case generates only an active system error.
///85: BDS_ISOBUS_RC_INV_FUNC_SEQU_DU16												Invalid execution sequence of function calls. Function |bds_isobus_setCaAddr| must be called before |bds_isobus_initComm|.
///
///==================================================================		   			===================================================================================================
///
///=======
///Code Example:
///=======
///============================================================================
///
///This Api should be called only once in application.
///
///PROGRAM Isobus_prg
///
///VAR
///
///    Flag_u8:USINT:=0;
///
///    EcuType_as8: ARRAY[1..20] OF STRING := ['Main ECU'];
///
///    EcuManu_as8: ARRAY[1..20] OF STRING := ['BOSCH REXROTH'];
///
///    ApplTask_as8: ARRAY[1..10] OF STRING := ['EHR'];    
///
///END_VAR
///
///(*call the api once*)
///
///IF(Flag_u8=0)THEN
///    
///    (* optionally define some ECU information of the controller application for the PGNs HW-ID and SW-ID: *)
///
///    bds_isobus_setCaInfo(2,16#0,ADR(EcuType_as8),ADR(EcuManu_as8),ADR(ApplTask_as8));
///        
///    (*define the controller application name, required for address claiming*)
///
///    bds_isobus_setCaName(1,16#00,16#02,16#00,16#01,16#81,16#01,16#01,16#33,BDS_ISOBUS_OWN_SN_DU32);
///    
///    (*define the initial source address and the CAN channel for the CA instance 1*)
///
///    bds_isobus_setCaAddr(1,BDS_CAN_3_D,16#10);
///    
///    (*initialize and start isobus communication for all instances on this CAN channel*)
///
///    bds_isobus_initComm(bds_can_Chnl_te.BDS_CAN_3_D, 50);
///    
///    Flag_u8:=1;
///    
///END_IF
///
///
///============================================================================
{attribute 'external_name' := 'cmp_rts_bds_isobus_setCaAddr'}
FUNCTION bds_isobus_setCaAddr : UINT
VAR_INPUT
	///ISOBUS instance number. This number identifies one instance of the ISOBUS stack.
	///
	///Value range: 1..n
	///n is the number of ISOBUS instances configured by easyConfig. 
	instanceNum_u8: USINT;
	///Indicates the CAN channel.
	///
	///Possible values for RC18-12/40, RC27-18/40:
	///   + BDS_CAN_1_D(0)
	///   + BDS_CAN_2_D(1)
	///   + BDS_CAN_3_D(2)
	///   + BDS_CAN_4_D(3)
	canChnl_e: bds_can_Chnl_te;
	///The own address, which is used as source address within all transmitted messages, until the address will be changed (e.g. by the service CommandedAddress).
	///A valid but already used source address leads only to an active system error. This behavior enables the application to use another source address. 
	///
	///Value range: 16#00 .. 16#FD.
	ownAddr_u8: USINT;
END_VAR

END_FUNCTION

// Communication API/ISOBUS/API/bds_isobus_getCaAddr
///This function reads the source address of one ISOBUS controller application.
///
///=======
/// Remarks:
///=======
///   + The source address which is read with this function is always the current address which is also used for the communication.
///   + The read source address may be the same as originally defined with the API function |bds_isobus_setCaAddr| but it does not have to be the same anymore.
///   + The CA (Controller Application) address may has been changed during run time
///	   + after the AddressClaiming procedure, if the arbitrary address capability feature is activated or
///	   + after a Commanded Address service call.
///   + The |GVL_isobus| is given for usage of defines.
///
///----------
/// FFI:
///----------
///This API can be used in trusted partitions only. See Freedom from Interference (FFI) concept for more details.
///
///==================================================================		  			===================================================================================================
///Return value    								  									Description
///==================================================================		  			===================================================================================================
///0..253																				Currently used CA address.
///254																					NullAddress, because function was executed with an error.
///
///==================================================================		   			===================================================================================================
///
///=======
///Code Example:
///=======
///============================================================================
///
///PROGRAM Isobus_prg
///
///VAR
///
///    Flag_u8:USINT:=0;
///
///    retval_u16: UINT;
///
///END_VAR
///
///(*call the api once*)
///
///IF(Flag_u8=0)THEN
///        
///    (*define the controller application name, required for address claiming*)
///
///    bds_isobus_setCaName(1,16#00,16#02,16#00,16#01,16#81,16#01,16#01,16#33,BDS_ISOBUS_OWN_SN_DU32);
///    
///    (*define the initial source address and the CAN channel for the CA instance 1*)
///
///    bds_isobus_setCaAddr(1,BDS_CAN_3_D,16#10);
///    
///    (*initialize and start isobus communication for all instances on this CAN channel*)
///
///    bds_isobus_initComm(bds_can_Chnl_te.BDS_CAN_3_D, 50);
///    
///    Flag_u8:=1;
///    
///END_IF
///
///(*get the actual address from the controller application instance 1*)
///
///retval_u16 := bds_isobus_getCaAddr(1);
///
///============================================================================
{attribute 'external_name' := 'cmp_rts_bds_isobus_getCaAddr'}
FUNCTION bds_isobus_getCaAddr : USINT
VAR_INPUT
	///ISOBUS instance number. This number identifies one instance of the ISOBUS stack.
	///
	///Value range: 1..n
	///n is the number of ISOBUS instances configured by easyConfig. 
	instanceNum_u8: USINT;
END_VAR

END_FUNCTION

// Communication API/ISOBUS/API/bds_isobus_getDiagnostic
///This function requests a DM1 or DM2 failure list from another controller application on another ECU.
///
///=======
/// Remarks:
///=======
///   + This function can be used by every instance of the ISOBUS communication stack to request a DM1 or DM2 failure list from another CA on other ECUs.
///   + This function can not be used to request a failure list from another CA on the own ECU.
///   + Before this function can be used, a corresponding failure list has to be defined with the function |bds_isobus_initDiagnostic|.
///   + The request of the DM1 failures with this function is not necessary, if the other controller sends the DM1 message cyclically.
///   + This function creates a PGN Request to the given destination address with the given DM type.
///   + The |GVL_isobus| is given for usage of defines.
///
///----------
/// FFI:
///----------
///This API can be used in trusted partitions only. See Freedom from Interference (FFI) concept for more details.
///
///==================================================================		  			===================================================================================================
///Return value    								  									Description
///==================================================================		  			===================================================================================================
///0: BDS_ISOBUS_RC_NO_ERRORS_DU16														Function was executed without errors.
///50: BDS_ISOBUS_RC_INV_ECU_ADDR_DU16													Invalid controller (ECU) address. Own CA address and 'null address' (16#FE) are not allowed.
///51: BDS_ISOBUS_RC_INV_DM_TYPE_DU16													Invalid DM failure type. Allowed values: BDS_ISOBUS_LIST_DM1_DU16 and BDS_ISOBUS_LIST_DM2_DU16
///80: BDS_ISOBUS_RC_INV_INST_NUM_DU16													Invalid instance number.
///
///==================================================================		   			===================================================================================================
///
///==================================================================		  			===================================================================================================
///dmType value	 								  									dmType Meaning
///==================================================================		  			===================================================================================================
///BDS_ISOBUS_LIST_DM1_DU16 (16#01)														DM1 failure list
///BDS_ISOBUS_LIST_DM2_DU16 (16#02)														DM2 failure list
///
///==================================================================		   			===================================================================================================
///

(*
=======
Code Example:
=======
============================================================================

VAR_GLOBAL
    (*allocate memory for DM1 failure list of another ECU*)
       isobus_dtcList1: bds_isobus_dtcList_ts;
END_VAR

PROGRAM Isobus_prg
VAR
    Flag_u8:USINT:=0;
    retval_u16: UINT;
    APPL_ISOBUS_INSTANCES_DU16: USINT:=10;
    isobus_appInst_as:ARRAY[1..10] OF bds_isobus_appInst_ts;
    ISOBUS_RX_BOXES_DU8: USINT:= 5;(* no of rx databoxes*)
    isobus_rxMsg_as: ARRAY[1..5] OF bds_isobus_rxMsg_ts; (*allocate memory for isobus rx databoxes*)
END_VAR

(*call the api once*)
IF(Flag_u8=0)THEN
    
    (*registers 10 isobus instances via the below bds_isobus_registerInstances api or by configuring it in easyConfig*)
   
    (*register isobus rx message boxes for instance 1 via bds_isobus_registerRxDataboxes api or via eC config*)
    
    (*init a DM1 failure list for instance 1 of the ECU with the address 77*)
   bds_isobus_initDiagnostic(1,  16#77, BDS_ISOBUS_LIST_DM1_DU16,ADR(gvl.isobus_dtcList1), 4,ADR(isobusDMCallback1));
    
    (*define the initial source address and the CAN channel for the CA instance 1*)
    bds_isobus_setCaAddr(1,BDS_CAN_3_D,16#10);
    
    (*initialize and start isobus communication for all instances on this CAN channel*)
    bds_isobus_initComm(bds_can_Chnl_te.BDS_CAN_3_D, 50);
    
    Flag_u8:=1;
    
END_IF

(*request the DM1 failure list from controller with address 77*)
 (*this is not required, if this controller sends the DM1 cyclically!*)

retval_u16:=bds_isobus_getDiagnostic(1, 16#77, BDS_ISOBUS_LIST_DM1_DU16);

(*the received DM1 failure list can be evaluated here*)


FUNCTION isobusDMCallback1
VAR
   isobus_nbrDtc_u16: UINT;
END_VAR

(*check the databox status and get the number of received DTCs*)

 IF (BDS_ISOBUS_BOXSTATUS_VALID_DU16 = bds_isobus_getRxDataboxStatus(1, 4, ADR(isobus_nbrDtc_u16))) THEN
   (*do anything*)
 END_IF
 
============================================================================
*)

{attribute 'external_name' := 'cmp_rts_bds_isobus_getDiagnostic'}
FUNCTION bds_isobus_getDiagnostic : UINT
VAR_INPUT
	///ISOBUS instance number. This number identifies one instance of the ISOBUS stack.
	///
	///Value range: 1..n
	///n is the number of ISOBUS instances configured by easyConfig. 
	instanceNum_u8: USINT;
	///Address of this controller application from which the DM1/DM2 failure list has to be received.
	///
	///Value range: 0..253, 255 (=all), own address is not allowed  
	destAddr_u8: USINT;
	///Type of the failure list (DM1/DM2) which is to be received. Optionally the conversion method version can be given, which is to be used in case of a received CM-Bit = 1.
	///
	///DTCs which are received with CM = 0 are always converted with conversion method version 4.
	dmType_u16: UINT;
END_VAR

// Communication API/ISOBUS/API/bds_isobus_initDiagnostic
///This function initializes a DM1 or DM2 failure list for the reception of these failures from other controllers and enables the reception of the corresponding DM1 or DM2 messages.
///
///=======
/// Remarks:
///=======
///   + This function must be called once per instance for the initialization of every failure type (DM1 or DM2) of each other controller, if the corresponding failures shall to be received.
///   + Every initialized failure list requires also a ISOBUS RX databox. It has to be taken into account during the configuration of the receive databoxes with easyConfig tool. These databoxes MUST NOT be initialized any more with the function |bds_isobus_initRxDatabox|.
///   + After the initialization of a failure list with this function, the corresponding data can be requested with the function |bds_isobus_getDiagnostic| and/or cyclic DM1/2 message will be received.
///   + After the reception of the whole DM1 message, the data will be converted in the following way:
///	   + The application can access the single DTCs using the structure elements of |bds_isobus_dtcList_ts|. (e.g. the PGN of the first DTC can be read directly with: isobus_dtcList1_s.dtc_as[0].spn_u32)
///	   + The function |bds_isobus_getRxDataboxStatus| returns directly the number of received DTCs as message length.
///	   + PGNs with format version 4 (CM = 0) and format versions 1..3 (CM = 1) are supported.
///	   + The received CM-Bit determines the used conversion method version. CM=0: always version 4 is used, CM=1: used version (1..3) is dependent on the parameter dmType_u16.  
///   + The DM1/DM2 DTC lists are limited to a size of 20 failures which can be received from other ECUs. Nevertheless DM1/DM2 messages with up to 29 failures can be received but during conversion the list will be truncated to the first 20 failures.
///   + This function internally initializes the given databox number for the reception and automatic conversion of DM1/DM2 failures. If the automatic conversion shall not be used the DM1/DM2 RX databox can be initialized as an alternative with the function |bds_isobus_initRxDatabox|. Then the databox contains the received raw data of the DM1/2 message which has to be interpreted accordingly by the application.
///   + The |GVL_isobus| is given for usage of defines.
///
///----------
/// FFI:
///----------
///This API can be used in trusted partitions only. See Freedom from Interference (FFI) concept for more details.
///
///==================================================================		  			===================================================================================================
///Return value    								  									Description
///==================================================================		  			===================================================================================================
///0: BDS_ISOBUS_RC_NO_ERRORS_DU16														Function was executed without errors.
///1: BDS_ISOBUS_RC_INVALID_ADDR_DU16													Address to data structure is Invalid.
///2: BDS_ISOBUS_RC_INV_DATABOX_DU16													Invalid databox number.
///20: BDS_ISOBUS_RC_PGN_SRC_EXIST_DU16												Another message box with the same PGN and source address is already defined.
///50: BDS_ISOBUS_RC_INV_ECU_ADDR_DU16													Invalid controller (ECU) address.
///51: BDS_ISOBUS_RC_INV_DM_TYPE_DU16													Invalid DM failure type. Allowed values: BDS_ISOBUS_LIST_DM1_DU16 and BDS_ISOBUS_LIST_DM2_DU16
///80: BDS_ISOBUS_RC_INV_INST_NUM_DU16													Invalid instance number.
///
///==================================================================		   			===================================================================================================
///
///==================================================================		  			===================================================================================================
///dmType value	 								  									dmType Meaning
///==================================================================		  			===================================================================================================
///BDS_ISOBUS_LIST_DM1_DU16 (16#01)														DM1 failure list, use CM version 3 for CM-Bit=1
///BDS_ISOBUS_LIST_DM2_DU16 (16#02)														DM2 failure list, use CM version 3 for CM-Bit=1
///BDS_ISOBUS_LIST_DM1_V1_DU16 (16#11)													DM1 failure list, use CM version 1 for CM-Bit=1
///BDS_ISOBUS_LIST_DM2_V1_DU16 (16#12)													DM2 failure list, use CM version 1 for CM-Bit=1
///BDS_ISOBUS_LIST_DM1_V2_DU16 (16#21)													DM1 failure list, use CM version 2 for CM-Bit=1
///BDS_ISOBUS_LIST_DM2_V2_DU16 (16#22)													DM2 failure list, use CM version 2 for CM-Bit=1
///BDS_ISOBUS_LIST_DM1_V3_DU16 (16#31)													DM1 failure list, use CM version 3 for CM-Bit=1
///BDS_ISOBUS_LIST_DM2_V3_DU16 (16#32)													DM2 failure list, use CM version 3 for CM-Bit=1
///
///==================================================================		   			===================================================================================================

(*
=======
Code Example:
=======
============================================================================

This Api should be called only once in application.

VAR_GLOBAL
    (*allocate memory for DM1 failure list of another ECU*)
	isobus_dtcList1: bds_isobus_dtcList_ts;
END_VAR

PROGRAM Isobus_prg
VAR
    Flag_u8:USINT:=0;
    retval_u16: UINT;
    APPL_ISOBUS_INSTANCES_DU16: USINT:=10;
    isobus_appInst_as:ARRAY[1..10] OF bds_isobus_appInst_ts;
    ISOBUS_RX_BOXES_DU8: USINT:= 5;(* no of rx databoxes*)
    isobus_rxMsg_as: ARRAY[1..5] OF bds_isobus_rxMsg_ts; (*allocate memory for isobus rx databoxes*)
END_VAR

(*call the api once*)
IF(Flag_u8=0)THEN
    
    (*registers 10 isobus instances via the below bds_isobus_registerInstances api or by configuring it in easyConfig*)
   
    (*register isobus rx message boxes for instance 1 via bds_isobus_registerRxDataboxes api or via eC config*)
    
    (*init a DM1 failure list for instance 1 of the ECU with the address 77*)
    retval_u16:=bds_isobus_initDiagnostic(1,  16#77, BDS_ISOBUS_LIST_DM1_DU16,ADR(gvl.isobus_dtcList1), 4,ADR(isobusDMCallback1));
    
    (*define the initial source address and the CAN channel for the CA instance 1*)
    bds_isobus_setCaAddr(1,BDS_CAN_3_D,16#10);
    
    (*initialize and start isobus communication for all instances on this CAN channel*)
    bds_isobus_initComm(bds_can_Chnl_te.BDS_CAN_3_D, 50);
    
    Flag_u8:=1;
    
END_IF


(*the received DM1 failure list can be evaluated here*)
FUNCTION isobusDMCallback1
VAR
    isobus_nbrDtc_u16: UINT;
END_VAR

(*check the databox status and get the number of received DTCs*)

 IF (BDS_ISOBUS_BOXSTATUS_VALID_DU16 = bds_isobus_getRxDataboxStatus(1, 4, ADR(isobus_nbrDtc_u16))) THEN
   (*do anything*)
 END_IF
 
============================================================================
*)
{attribute 'external_name' := 'cmp_rts_bds_isobus_initDiagnostic'}
FUNCTION bds_isobus_initDiagnostic : UINT
VAR_INPUT
	///ISOBUS instance number. This number identifies one instance of the ISOBUS stack.
	///
	///Value range: 1..n
	///n is the number of ISOBUS instances configured by easyConfig. 
	instanceNum_u8: USINT;
	///Address of this controller application from which the DM1/DM2 failure list has to be received.
	///
	///Value range: 0..253 
	srcAddr_u8: USINT;
	///Type of the failure list (DM1/DM2) which is to be received. Optionally the conversion method version can be given, which is to be used in case of a received CM-Bit = 1.
	///
	///DTCs which are received with CM = 0 are always converted with conversion method version 4.
	dmType_u16: UINT;
	///Pointer to a DM1/DM2 failure list, which has to be defined by the application.
	///
	///Pointer to a variable of data type bds_isobus_dtcList_ts.
	dtcList_ps: POINTER TO bds_isobus_dtcList_ts;
	///The number of a ISOBUS receive databox, which can be exclusively used for receiving of the DM1/2 message. This databox MUST NOT be initialized additionally with the function |bds_isobus_initRxDatabox|.
	///
	///Value range: 1..n
	///n is the number of receive databoxes configured by easyConfig or alternatively with function |bds_isobus_registerRxDataboxes|. 
	boxNum_u16: UINT;
	///Pointer to a callback function of data type UINT which is called after a new message was received completely. The execution time of the callback function should be short to be able to meet the time conditions within the ISOBUS stack. 
	func_pf: POINTER TO BOOL;
END_VAR

// Communication API/ISOBUS/API/bds_isobus_initRxDatabox
///This function initializes a ISOBUS receive databox. The ISOBUS messages can be received only with ISOBUS receive databoxes.
///
///=======
/// Remarks:
///=======
///   + This function must be called during the configuration of the ISOBUS communication stack once for each ISOBUS receive message.
///   + Before the RX databoxes can be initialized with this function, the required number of receive databoxes has to be configured first with easyConfig tool or alternatively with function |bds_isobus_registerRxDataboxes|.
///   + Each ISOBUS RX databox requires an own data array or a data structure. The pointer to this data field is required for the initialization of a ISOBUS receive databox. The received data then will be stored in this data field.
///   + The data array for the received data may have a length of more than 8 bytes (see parameter description below). 
///   + The execution time of the callback function should be short to be able to meet the time conditions within the ISOBUS stack.
///   + If the same CAN bus is also used for further communication, ensure that the CAN IDs are uniquely assigned.
///   + The meaning of this function is similar to the system function |bds_can_initRxDatabox|.
///   + In addition to the ISOBUS specifications, this function can be used for the reception of ISOBUS single frame PDU1 format messages which are sent to the own network adddress as well as to other destination addresses.
///   + The definition of a destination address within PDU1 format PGNs is mandatory.
///   + Important(Non Standard PGN): For the reception of PDU1 format messages to the own network address the PDU Specific part (=Destination) of the PGN should be defined with the NULL address value (=16#FE) instead of the own address. Otherwise the own address within the RX databoxes may not match any more with the real own address after an address claiming.
///   + Important(Standard PGN):To Receive the Data of PGN's like Address Claim,Request PGN,Name Management and Stop start(DM13)  which are sent to the own network adddress (PDU Specific part =16#FF) or   (PDU Specific part=Destination) can be received by registering the Databox with the respective PGN. PGN Data will be consumed and processed by the ISOBUS Stack but Data will be available for application.
///   + Example: Application has to receive Address Claimed PGN (16#EE00) data and it is also applicable for Request PGN,Name Management and Stop start(DM13)(Standard  PGN)
///   + The |GVL_isobus| is given for usage of defines.
///
///----------
/// FFI:
///----------
///This API can be used in trusted partitions only. See Freedom from Interference (FFI) concept for more details.
///
///==================================================================		  			===================================================================================================
///Return value    								  									Description
///==================================================================		  			===================================================================================================
///0: BDS_ISOBUS_RC_NO_ERRORS_DU16														Function was executed without errors.
///2: BDS_ISOBUS_RC_INV_DATABOX_DU16													Invalid databox number.
///3: BDS_ISOBUS_RC_INV_PGN_DU16														Invalid parameter group number (PGN).
///4 BDS_ISOBUS_RC_INV_SRC_DU16														Invalid source address.
///5: BDS_ISOBUS_RC_INV_TIMEOUT_DU16													Invalid timeout value.
///6: BDS_ISOBUS_RC_INV_DATA_LEN_DU16													Invalid data length.
///7:BDS_ISOBUS_RC_INV_DATA_PTR_DU16													Invalid address pointer.
///9:BDS_ISOBUS_RC_INV_STARTTIMEOUT_DU16												Invalid start timeout value.
///20: BDS_ISOBUS_RC_PGN_SRC_EXIST_DU16												Another message box with the same PGN and source address is alraedy defined.
///80: BDS_ISOBUS_RC_INV_INST_NUM_DU16													Invalid instance number.
///86: BDS_ISOBUS_RC_PGN_USED_INTERNAL_DU16											Registered PGN Data will be consumed by ISOBUS Stack.Data will be available for the application after  ISOBUS Stack processing
///
///==================================================================		   			===================================================================================================
///
///==================================================================		  			===================================================================================================
///Standard PGN	 								  									Data in Databox
///==================================================================		  			===================================================================================================
///Registered as "16#EEFF"																Receives only data which is broadcasted(PDU Specific part =16#FF).ex: bds_isobus_initRxDatabox(1, 02, 16#EEFF,  16#01, 1000, 5000, 25,msgRx3Data_au8, 0);It only receives the data which is brodcasted from source address 16#01.
///Registered "16#EE<own address>"														Receives data which is directed to the ECU by its own address (PDU Specific part=Destination).ex: bds_isobus_initRxDatabox(1, 02, 16#EE04,  16#01, 1000, 5000, 25,msgRx3Data_au8, 0);It only receives the data which is directed to the ECU by requesting with its own address(16#04).Note:If you initialize Databox with "16#EEFE" you only receive data with whose PDU Specific part is Null(16#FE).
///
///==================================================================		   			===================================================================================================
///
///=======
///Code Example:
///=======
///============================================================================
///
///This Api should be called only once in application.
///
///VAR_GLOBAL
///
///    (*global data buffer for isobus Rx message*)
///
///    msgRx2Data_au8: ARRAY[1..8] OF USINT;
///
///END_VAR
///
///PROGRAM Isobus_prg
///
///VAR
///
///    Flag_u8:USINT:=0;
///
///    retval_u16: UINT;
///
///    APPL_ISOBUS_INSTANCES_DU16: USINT:=10;
///
///    isobus_appInst_as:ARRAY[1..10] OF bds_isobus_appInst_ts;
///
///    ISOBUS_RX_BOXES_DU8: USINT:= 5;(* no of rx databoxes*)
///
///    isobus_rxMsg_as: ARRAY[1..5] OF bds_isobus_rxMsg_ts; (*allocate memory for isobus rx databoxes*)
///
///END_VAR
///
///(*call the api once*)
///
///IF(Flag_u8=0)THEN
///    
///    (*registers 10 isobus instances via the below api or by configuring it in easyConfig*)
///
///    bds_isobus_registerInstances(ADR(isobus_appInst_as), APPL_ISOBUS_INSTANCES_DU16);
///    
///    (*register isobus rx message boxes for instance 1*)
///
///    bds_isobus_registerRxDataboxes(1,ADR(isobus_rxMsg_as),ISOBUS_RX_BOXES_DU8);
///    
///    (*initalize rx databox messages for databox 1 of instance 1 with pgn 16#7789*)
///
///    retval_u16:= bds_isobus_initRxDatabox(1, 1, 16#7789, 16#04, 2000, 6000, 8,ADR(gvl.msgRx2Data_au8),ADR(Rxcallback));
///    
///    (*define the controller application name, required for address claiming*)
///
///    bds_isobus_setCaName(1,16#00,16#02,16#00,16#01,16#81,16#01,16#01,16#33,BDS_ISOBUS_OWN_SN_DU32);
///    
///    (*define the initial source address and the CAN channel for the CA instance 1*)
///
///    bds_isobus_setCaAddr(1,BDS_CAN_3_D,16#10);
///    
///    (*initialize and start isobus communication for all instances on this CAN channel*)
///
///    bds_isobus_initComm(bds_can_Chnl_te.BDS_CAN_3_D, 50);
///    
///    Flag_u8:=1;
///    
///END_IF
///
///FUNCTION Rxcallback
///
///VAR
///
///END_VAR
///
///(*The received message is further sent on can for verification*)
///
///bds_can_SendData(bds_can_Chnl_te.BDS_CAN_3_D,16#CB3,1,8,ADR(gvl.msgRx2Data_au8));
///============================================================================
{attribute 'external_name' := 'cmp_rts_bds_isobus_initRxDatabox'}
FUNCTION bds_isobus_initRxDatabox : UINT
VAR_INPUT
	///ISOBUS instance number. This number identifies one instance of the ISOBUS stack.
	///
	///Value range: 1..n
	///n is the number of ISOBUS instances configured by easyConfig. 
	instanceNum_u8: USINT;
	///Number of a ISOBUS receive databox.
	///
	///Value range: 1..n
	///n is the number of receive databoxes configured by easyConfig or alternatively with function |bds_isobus_registerRxDataboxes|.
	boxNum_u16: UINT;
	///Parameter group number (PGN) of the message to be received with this databox. For PDU1 format PGNs see remark above.
	///
	///Value range: 0..16#3FFFF (18 bit) 
	pgn_u32: UDINT;
	///Source address of the transmitter of the ISOBUS message from which the message has to be received.
	///
	///Value range: 16#00..16#FD 
	src_u8: USINT;
	///With this time (in ms) the cyclic reception of this message can be supervised. If a cyclic message was not received during this time, then the RX databox status will be set to ISOBUS_BOXSTATUS_INV_TIMEOUT_DU16. This time is only applicable after the first reception of this ISOBUS message after the initialization. 
	timeout_u16: UINT;
	///With this time (in ms) the first reception of this message can be supervised. If a first message after initialization was not received during this time, then the RX databox status will be set to ISOBUS_BOXSTATUS_INV_TIMEOUT_DU16. This time is only applicable for the first time after the (re-)initialization. 
	///
	///Value range: 10..65000 [ms] or 0 = no time supervision  
	startTimeout_u16: UINT;
	///Size of the data array/structure below. A ISOBUS message may consist of several single CAN messages, if the number of data bytes is more than 8.
	///
	///Value range: 1..117440512
	lenMax_u32: UDINT;
	///Pointer to a data array or a data structure, in which the received data can be stored. The size of this array/structure has to be given within the previous parameter (lenMax_u32).
	///
	///It is neccessary to declare the buffer array/structure as a global variable!
	data_pau8: POINTER TO USINT;
	///Pointer to a callback function of datatype UINT which is called after a new message was received completely. The execution time of the callback function should be short to be able to meet the time conditions within the ISOBUS stack.Function must be coded within the application program.
	///Optional a NULL pointer can be assigned to disable the callback function.
	func_pf: POINTER TO BOOL;
END_VAR

END_FUNCTION

// Communication API/ISOBUS/API/bds_isobus_registerRxDataboxes
///This function registers memory for ISOBUS receive databoxes and therefore defines the maximal number of usable ISOBUS receive databoxes per instance.
///
///=======
/// Remarks:
///=======
///   + This function must be called once during the configuration of the ISOBUS communication stack before |bds_isobus_initComm|.
///   + After the execution of this function, each ISOBUS receive databox has to be initialized with |bds_isobus_initRxDatabox| before using.
///   + The |GVL_isobus| is given for usage of defines.
///   + This function should be called only once in the application.
///   
///----------
/// Notice:
///----------
///
///This API-function can be used alternatively to the ISOBUS configuration with easyConfig. If this function is used, then the number of ISOBUS RX databoxes is to be configured to 0 in easyConfig.
///
///----------
/// FFI:
///----------
///This API can be used in trusted partitions only. See Freedom from Interference (FFI) concept for more details.
///
///==================================================================		  			===================================================================================================
///Return value    								  									Description
///==================================================================		  			===================================================================================================
///0: BDS_ISOBUS_RC_NO_ERRORS_DU16														Function was executed without errors.
///1: BDS_ISOBUS_RC_INVALID_ADDR_DU16													Address to data array is Invalid.
///8: BDS_ISOBUS_RC_OVERLAP_ADDR_DU16													Address overlaps with an already existing buffer.
///22: BDS_ISOBUS_RC_CFG_NOTALLOWED_DU16												Function must be called before bds_isobus_initComm, but it was called afterwards.
///80: BDS_ISOBUS_RC_INV_INST_NUM_DU16													Invalid instance number.
///
///==================================================================		   			===================================================================================================
///
///=======
///Code Example:
///=======
///============================================================================
///
///This Api should be called only once in application.
///
/// 
///PROGRAM Isobus_prg
///
///VAR
///
///    Flag_u8:USINT:=0;
///
///    retval_u16: UINT;
///
///    isobus_appInst_as:ARRAY[1..10] OF bds_isobus_appInst_ts;
///
///    ISOBUS_RX_BOXES_DU8: USINT:= 5;(* no of rx databoxes*)
///
///    APPL_ISOBUS_INSTANCES_DU16: USINT:=10;
///
///    isobus_rxMsg_as: ARRAY[1..5] OF bds_isobus_rxMsg_ts; (*allocate memory for isobus rx databoxes*)
///
///END_VAR
///
///(*call the api once*)
///
///IF(Flag_u8=0)THEN
///    
///    (*registers 10 isobus instances*)
///
///    bds_isobus_registerInstances(ADR(isobus_appInst_as), APPL_ISOBUS_INSTANCES_DU16);
///    
///    (*register isobus rx message boxes for instance 1*)
///
///    retval_u16:=bds_isobus_registerRxDataboxes(1,ADR(isobus_rxMsg_as),ISOBUS_RX_BOXES_DU8);
///    
///    Flag_u8:=1;
///    
///END_IF
///
///
///============================================================================
{attribute 'external_name' := 'cmp_rts_bds_isobus_registerRxDataboxes'}
FUNCTION bds_isobus_registerRxDataboxes : UINT
VAR_INPUT
	///ISOBUS instance number. This number identifies one instance of the ISOBUS stack.
	///
	///Value range: 1..n
	///n is the number of ISOBUS instances configured by easyConfig. 
	instanceNum_u8: USINT;
	///Pointer to an array of data type bds_isobus_rxMsg_ts.
	///
	///Note:
	///The buffer will be managed by the BSW. The application has only to declare the buffer (memory space).
	///It is necessary to declare the buffer array as a global variable! 
	mem_pas: POINTER TO bds_isobus_rxMsg_ts;
	///Size of the array above, which corresponds to the number of usable isobus receive databoxes. 
	num_u16: UINT;
END_VAR

END_FUNCTION

// Communication API/ISOBUS/API/bds_isobus_registerInstances
///This function registers memory for all required ISOBUS controller application instances (CA) and therefore defines the maximal number of usable CA instances.
///
///=======
/// Remarks:
///=======
///   + This function stores the pointer to an array of the data memory structure which can be used by the ISOBUS instances and the size of this array.
///   + This function shall be called internally during ISOBUS module initialization. The registered memory size depends on the configuration within easyConfig.
///   + The |GVL_isobus| is given for usage of defines.
///
///----------
/// WARNING:
///----------
///
///This function should be called only once in the application.
///
///----------
/// FFI:
///----------
///This API can be used in trusted partitions only. See Freedom from Interference (FFI) concept for more details.
///
///==================================================================		  			===================================================================================================
///Return value    								  									Description
///==================================================================		  			===================================================================================================
///0: BDS_ISOBUS_RC_NO_ERRORS_DU16														Function was executed without errors.
///1: BDS_ISOBUS_RC_INVALID_ADDR_DU16													Invalid address to the data array.
///8: BDS_ISOBUS_RC_OVERLAP_ADDR_DU16													Address overlaps with other buffers.
///80: BDS_ISOBUS_RC_INV_INST_NUM_DU16													Invalid CA instance number.
///84: BDS_ISOBUS_RC_REGINST_NOT_ALLOWED_DU16											Function call is not allowed outside OsIniProc().
///
///==================================================================		   			===================================================================================================
///
///=======
///Code Example:
///=======
///============================================================================
///
///This Api should be called only once in application.
/// 
///PROGRAM Isobus_prg
///
///VAR
///    Flag_u8:USINT:=0;
///
///    retval_u16: UINT;
///
///    isobus_appInst_as:ARRAY[1..10] OF bds_isobus_appInst_ts;
///
///    APPL_ISOBUS_INSTANCES_DU16: USINT:=10;
///
///END_VAR
///
///(*call the api once*)
///
///IF(Flag_u8=0)THEN
///    
///    (*registers 10 isobus instances*)
///
///    retval_u16:=bds_isobus_registerInstances(ADR(isobus_appInst_as), APPL_ISOBUS_INSTANCES_DU16);
///
///    Flag_u8:=1;
///    
///END_IF
///
///============================================================================
{attribute 'external_name' := 'cmp_rts_bds_isobus_registerInstances'}
FUNCTION bds_isobus_registerInstances : UINT
VAR_INPUT
	///Pointer to data memory array of all instances
	mem_pas: POINTER TO bds_isobus_appInst_ts;
	///Size of the array above, which corresponds to the number of usable ISOBUS controller application instances.
	///
	///Value range: 1..10
	num_u16: UINT;
END_VAR

END_FUNCTION

